Yaskawa INFORM job: SPLITTE3.JBI

/JOB
//NAME SPLITTE3
//POS
///NPOS 15,0,0,0,0,0
///TOOL 1
///POSTYPE PULSE
///PULSE
C00000=14,20,-5,30,-45,60
C00001=18,24,-10,30,-45,60
C00002=14,20,-5,30,-45,60
C00003=18,24,-10,30,-45,60
C00004=14,20,-5,30,-45,60
C00005=18,24,-10,30,-45,60
C00006=14,20,-5,30,-45,60
C00007=18,24,-10,30,-45,60
C00008=14,20,-5,30,-45,60
C00009=18,24,-10,30,-45,60
C00010=14,20,-5,30,-45,60
C00011=18,24,-10,30,-45,60
C00012=14,20,-5,30,-45,60
C00013=18,24,-10,30,-45,60
C00014=14,20,-5,30,-45,60
//INST
///DATE 2026/10/26 01:19
///COMM Generated using RoboDK
///ATTR SC,RW
///GROUP1 RB1
NOP
MOVL C00000 V=200.0
MOVL C00001 V=200.0
MOVL C00002 V=200.0
MOVL C00003 V=200.0
MOVL C00004 V=200.0
MOVL C00005 V=200.0
MOVL C00006 V=200.0
MOVL C00007 V=200.0
MOVL C00008 V=200.0
MOVL C00009 V=200.0
MOVL C00010 V=200.0
MOVL C00011 V=200.0
MOVL C00012 V=200.0
MOVL C00013 V=200.0
MOVL C00014 V=200.0
END
